FUNCTION "FC_StlNoPar" : Void
{ S7_Optimized_Access := 'FALSE' ; S7_Pass_Registers := 'TRUE' }
VERSION : 0.1

BEGIN
NETWORK
TITLE =
      NOP 0;
END_FUNCTION

